// TIA Portal V20 export
Screen "190RB06_V23"  1276x673
  ScreenItem "Graphic view_1" at 181,100 size 790x526  Type=HmiGraphicView
  ScreenItem "Line_Header_X0_Y64" at 0,64 size 1276x0  Type=HmiLine
  ScreenItem "permanentareaborderrectangle" at 0,0 size 0x0  Type=HmiRectangle
  ScreenItem "Button_Back" at 2,2 size 90x60  Type=HmiButton
  ScreenItem "Title_ScreenOverview_X390_Y2_2" at 392,4 size 510x57  Type=HmiTextBox
  ScreenItem "Fusszeile_Button_ManualOPMode1_4" at 1181,2 size 90x60  Type=HmiButton
  ScreenItem "Title_ScreenOverview_X390_Y2_1" at 1130,78 size 139x57  Type=HmiTextBox
  ScreenItem "Title_ScreenOverview_X390_Y2_3" at 1130,144 size 139x57  Type=HmiTextBox
  ScreenItem "Title_ScreenOverview_X390_Y2_4" at 1130,144 size 139x57  Type=HmiTextBox
  ScreenItem "文本域_19" at 964,95 size 134x40  Type=HmiTextBox
  ScreenItem "Line_19" at 911,143 size 68x20  Type=HmiLine
  ScreenItem "Line_2" at 891,245 size 132x1  Type=HmiLine
  ScreenItem "文本域_4" at 1047,300 size 134x40  Type=HmiTextBox
  ScreenItem "Line_5" at 887,316 size 160x47  Type=HmiLine
  ScreenItem "Line_3" at 897,421 size 142x12  Type=HmiLine
  ScreenItem "文本域_5" at 1023,543 size 134x40  Type=HmiTextBox
  ScreenItem "Line_6" at 911,560 size 104x13  Type=HmiLine
  ScreenItem "Line_11" at 700,385 size 27x87  Type=HmiLine
  ScreenItem "文本域_6" at 632,582 size 134x40  Type=HmiTextBox
  ScreenItem "Line_7" at 594,569 size 33x36  Type=HmiLine
  ScreenItem "文本域_1" at 435,509 size 134x40  Type=HmiTextBox
  ScreenItem "Line_1" at 515,478 size 15x26  Type=HmiLine
  ScreenItem "文本域_7" at 319,582 size 134x40  Type=HmiTextBox
  ScreenItem "Line_4" at 377,542 size 22x35  Type=HmiLine
  ScreenItem "Line_8" at 192,566 size 73x27  Type=HmiLine
  ScreenItem "文本域_8" at 47,583 size 134x40  Type=HmiTextBox
  ScreenItem "Line_9" at 193,472 size 74x19  Type=HmiLine
  ScreenItem "文本域_11" at 18,374 size 134x40  Type=HmiTextBox
  ScreenItem "Line_10" at 157,361 size 90x38  Type=HmiLine
  ScreenItem "Line_12" at 191,226 size 81x98  Type=HmiLine
  ScreenItem "文本域_16" at 13,95 size 134x40  Type=HmiTextBox
  ScreenItem "Line_15" at 153,127 size 92x25  Type=HmiLine
  ScreenItem "Line_17" at 399,252 size 41x91  Type=HmiLine
  ScreenItem "Line_20" at 434,109 size 99x140  Type=HmiLine
  ScreenItem "文本域_20" at 300,68 size 134x40  Type=HmiTextBox
  ScreenItem "文本域_13" at 453,69 size 134x40  Type=HmiTextBox
  ScreenItem "Line_13" at 548,117 size 26x30  Type=HmiLine
  ScreenItem "文本域_14" at 653,81 size 134x40  Type=HmiTextBox
  ScreenItem "Line_14" at 755,134 size 10x48  Type=HmiLine
  ScreenItem "Title_ScreenOverview_X390_Y2_44" at 338,111 size 52x19  Type=HmiTextBox
  ScreenItem "Title_ScreenOverview_X390_Y2_45" at 338,131 size 25x21  Type=HmiTextBox
  ScreenItem "Title_ScreenOverview_X390_Y2_46" at 365,131 size 25x21  Type=HmiTextBox
  ScreenItem "Title_ScreenOverview_X390_Y2_5" at 487,108 size 52x19  Type=HmiTextBox
  ScreenItem "Title_ScreenOverview_X390_Y2_6" at 487,128 size 25x21  Type=HmiTextBox
  ScreenItem "Title_ScreenOverview_X390_Y2_7" at 514,128 size 25x21  Type=HmiTextBox
  ScreenItem "Title_ScreenOverview_X390_Y2_8" at 693,121 size 52x19  Type=HmiTextBox
  ScreenItem "Title_ScreenOverview_X390_Y2_9" at 693,141 size 25x21  Type=HmiTextBox
  ScreenItem "Title_ScreenOverview_X390_Y2_10" at 720,141 size 25x21  Type=HmiTextBox
  ScreenItem "Title_ScreenOverview_X390_Y2_11" at 1001,135 size 52x19  Type=HmiTextBox
  ScreenItem "Title_ScreenOverview_X390_Y2_12" at 1001,155 size 25x21  Type=HmiTextBox
  ScreenItem "Title_ScreenOverview_X390_Y2_13" at 1028,155 size 25x21  Type=HmiTextBox
  ScreenItem "Title_ScreenOverview_X390_Y2_14" at 1082,360 size 25x21  Type=HmiTextBox
  ScreenItem "Title_ScreenOverview_X390_Y2_15" at 1082,340 size 52x19  Type=HmiTextBox
  ScreenItem "Title_ScreenOverview_X390_Y2_16" at 1109,360 size 25x21  Type=HmiTextBox
  ScreenItem "Title_ScreenOverview_X390_Y2_17" at 1057,588 size 52x19  Type=HmiTextBox
  ScreenItem "Title_ScreenOverview_X390_Y2_18" at 1057,608 size 25x21  Type=HmiTextBox
  ScreenItem "Title_ScreenOverview_X390_Y2_19" at 1084,608 size 25x21  Type=HmiTextBox
  ScreenItem "Title_ScreenOverview_X390_Y2_20" at 675,622 size 52x19  Type=HmiTextBox
  ScreenItem "Title_ScreenOverview_X390_Y2_21" at 675,642 size 25x21  Type=HmiTextBox
  ScreenItem "Title_ScreenOverview_X390_Y2_22" at 702,642 size 25x21  Type=HmiTextBox
  ScreenItem "Title_ScreenOverview_X390_Y2_23" at 476,549 size 52x19  Type=HmiTextBox
  ScreenItem "Title_ScreenOverview_X390_Y2_24" at 476,569 size 25x21  Type=HmiTextBox
  ScreenItem "Title_ScreenOverview_X390_Y2_25" at 503,569 size 25x21  Type=HmiTextBox
  ScreenItem "Title_ScreenOverview_X390_Y2_26" at 365,622 size 52x19  Type=HmiTextBox
  ScreenItem "Title_ScreenOverview_X390_Y2_27" at 365,642 size 25x21  Type=HmiTextBox
  ScreenItem "Title_ScreenOverview_X390_Y2_28" at 392,642 size 25x21  Type=HmiTextBox
  ScreenItem "Title_ScreenOverview_X390_Y2_29" at 86,627 size 52x19  Type=HmiTextBox
  ScreenItem "Title_ScreenOverview_X390_Y2_30" at 86,647 size 25x21  Type=HmiTextBox
  ScreenItem "Title_ScreenOverview_X390_Y2_31" at 113,647 size 25x21  Type=HmiTextBox
  ScreenItem "Title_ScreenOverview_X390_Y2_32" at 58,414 size 52x19  Type=HmiTextBox
  ScreenItem "Title_ScreenOverview_X390_Y2_33" at 58,434 size 25x21  Type=HmiTextBox
  ScreenItem "Title_ScreenOverview_X390_Y2_34" at 85,434 size 25x21  Type=HmiTextBox
  ScreenItem "Title_ScreenOverview_X390_Y2_35" at 50,134 size 52x19  Type=HmiTextBox
  ScreenItem "Title_ScreenOverview_X390_Y2_36" at 77,154 size 25x21  Type=HmiTextBox
  ScreenItem "Title_ScreenOverview_X390_Y2_37" at 50,154 size 25x21  Type=HmiTextBox
  ScreenItem "Rectangle_1" at 0,0 size 131x48  Type=HmiRectangle
  ScreenItem "文本域_15" at 2,1 size 105x45  Type=HmiTextBox
  ScreenItem "圆_1" at 0,0 size 100x30  Type=HmiCircle
  ScreenItem "圆_2" at 0,0 size 100x30  Type=HmiCircle
  ScreenItem "Rectangle_13" at 0,0 size 165x48  Type=HmiRectangle
  ScreenItem "文本域_12" at 2,1 size 132x45  Type=HmiTextBox
  ScreenItem "圆_5" at 0,0 size 100x30  Type=HmiCircle
  ScreenItem "圆_6" at 0,0 size 100x30  Type=HmiCircle
  ScreenItem "Rectangle_2" at 0,0 size 165x48  Type=HmiRectangle
  ScreenItem "文本域_17" at 2,1 size 132x45  Type=HmiTextBox
  ScreenItem "圆_3" at 0,0 size 100x30  Type=HmiCircle
  ScreenItem "圆_4" at 0,0 size 100x30  Type=HmiCircle
  ScreenItem "Rectangle_3" at 0,0 size 165x48  Type=HmiRectangle
  ScreenItem "文本域_2" at 2,1 size 132x45  Type=HmiTextBox
  ScreenItem "圆_7" at 0,0 size 100x30  Type=HmiCircle
  ScreenItem "圆_8" at 0,0 size 100x30  Type=HmiCircle
  ScreenItem "Rectangle_4" at 0,0 size 165x48  Type=HmiRectangle
  ScreenItem "文本域_3" at 2,1 size 132x45  Type=HmiTextBox
  ScreenItem "圆_9" at 0,0 size 100x30  Type=HmiCircle
  ScreenItem "圆_10" at 0,0 size 100x30  Type=HmiCircle
  ScreenItem "Rectangle_5" at 0,0 size 131x48  Type=HmiRectangle
  ScreenItem "文本域_9" at 2,1 size 105x45  Type=HmiTextBox
  ScreenItem "圆_11" at 0,0 size 100x30  Type=HmiCircle
  ScreenItem "圆_12" at 0,0 size 100x30  Type=HmiCircle
